// TIA Portal V20 export
// export: Created 2026-10-19T18:38:08.4370459Z, ExportSetting WithDefaults, DisplayName Totally Integrated Automation Portal, DisplayVersion V20 Update 6, DisplayName TIA Portal Openness, DisplayVersion V20 Update 6, DisplayName TIA Portal Version Control Interface, DisplayVersion V20 Update 6, DisplayName SINAMICS Startdrive Advanced, DisplayVersion V20 SP1, DisplayName SINAMICS Startdrive G130, G150, S120, S150, SINAMICS MV, G220, S200, S210, DisplayVersion V20 SP1, DisplayName SINAMICS Startdrive G110M, G120, G120C, G120D, G120P, G115D, DisplayVersion V20 SP1, DisplayName STEP 7 Professional, DisplayVersion V20 Update 6, DisplayName STEP 7 Safety, DisplayVersion V20 Update 2, DisplayName WinCC Basic/Comfort/Advanced, DisplayVersion V20 Update 6, DisplayName WinCC Unified, DisplayVersion V20 Update 6
FUNCTION "ID_Decode_F" : Void   // FC3, SCL
{ S7_Optimized_Access := 'TRUE' }
VERSION : 0.1
// stored: AutoNumber true, IsIECCheckEnabled false, SetENOAutomatically false, UDAEnableTagReadback false
   VAR_INPUT
      ID : DInt;
   END_VAR
   VAR_IN_OUT
      ID_Decoded : "ID_Decoded";
   END_VAR
   VAR_TEMP
      Temp : UInt;
   END_VAR
BEGIN

   // Extract XX (first two digits)
   #ID_Decoded.Device_Type := #ID / 10000;        // 123456 / 10000 = 12

   // Extract YY (middle two digits)
   #ID_Decoded.Level := (#ID MOD 10000) / 100; // 123456 % 10000 = 3456 → 3456 / 100 = 34

   // Extract ZZ (last two digits)
   #ID_Decoded.VTD := #ID MOD 100;       // 123456 % 100 = 56
END_FUNCTION
